Fanuc KAREL source: kt00193.KL

-- PROVISIONAL review KL for V940-1; original PC SHA256 349e2b4faf9e85752dfdc52194297034923c2caf5873f7ec9537f37942569fc1
-- Incomplete behavior may be omitted. Consult companion uncertainty JSON. Do not deploy.
PROGRAM KT00193
%NOLOCKGROUP
VAR
  B1 : BOOLEAN
  B2 : BOOLEAN
  OUT : BOOLEAN
BEGIN
  B1 = TRUE
  B2 = FALSE
  B1 = TRUE
  B2 = FALSE
  OUT = (B1 AND B2)
END KT00193
